FUNCTION_BLOCK FB_JamConveyor EXTENDS FB_ConveyorBase
VAR
    jamTimer : TON;
END_VAR

METHOD PROTECTED DetectJam : BOOL
VAR_INPUT
    blocked : BOOL;
END_VAR
jamTimer(IN := blocked, PT := T#300ms);
DetectJam := jamTimer.Q;
END_METHOD

END_FUNCTION_BLOCK

(* stored: Version 1.1.0.1, ProductVersion 3.1 *)
